FUNCTION_BLOCK FB_Snapshot		// 이번 스캔의 장비 상태를 한 번에 복사. 이후 단계는 이 사본만 읽는다
VAR_IN_OUT
	iq_aipPcs		: ARRAY[1..GVL_PARAM.PCS_COUNT] OF I_Pcs;
	iq_aipBms		: ARRAY[1..GVL_PARAM.BMS_COUNT] OF I_Bms;
	iq_aipMeter		: ARRAY[1..GVL_PARAM.METER_COUNT] OF I_Meter;
END_VAR
VAR_IN_OUT CONSTANT
	iq_astUnitCfg	: ARRAY[1..GVL_PARAM.UNIT_COUNT] OF ST_UnitCfg;
END_VAR
VAR_OUTPUT
	q_astUnit		: ARRAY[1..GVL_PARAM.UNIT_COUNT] OF ST_UnitState;
	q_astBms		: ARRAY[1..GVL_PARAM.BMS_COUNT] OF ST_BatState;
	q_astMeter		: ARRAY[1..GVL_PARAM.METER_COUNT] OF ST_MeterState;
END_VAR
VAR_TEMP
	i				: UINT;
	nPcs			: UINT;
	stNoUnit		: ST_UnitState;		// 빈 칸: 통신 없음, 상태 Unknown
	stNoBms			: ST_BatState;
	stNoMeter		: ST_MeterState;
	k				: UINT;		// [결함 9 수정 2026-11-03: 추가]
END_VAR

// 유닛: 구성표의 PCS 번호·PCS 안 번호로 찾음
FOR i := 1 TO GVL_PARAM.UNIT_COUNT DO
	nPcs := iq_astUnitCfg[i].nPcs;
	IF nPcs >= 1 AND nPcs <= GVL_PARAM.PCS_COUNT AND_THEN iq_aipPcs[nPcs] <> 0 THEN
		q_astUnit[i] := iq_aipPcs[nPcs].M_GetUnitState(iq_astUnitCfg[i].nSub);
		q_astUnit[i].stP := M_FixVal(q_astUnit[i].stP);	// [결함 9 수정 2026-11-03: NaN·무한대 → 0·무효]
		q_astUnit[i].stQ := M_FixVal(q_astUnit[i].stQ);
	ELSE
		q_astUnit[i] := stNoUnit;
	END_IF
END_FOR

FOR i := 1 TO GVL_PARAM.BMS_COUNT DO
	IF iq_aipBms[i] <> 0 THEN
		q_astBms[i] := iq_aipBms[i].BatState;
		q_astBms[i].stSoc := M_FixVal(q_astBms[i].stSoc);	// [결함 9 수정 2026-11-03: NaN·무한대 → 0·무효, 한도는 0]
		q_astBms[i].stSoh := M_FixVal(q_astBms[i].stSoh);
		IF NOT F_CmdOk(q_astBms[i].fPChgMax, 0.0) THEN q_astBms[i].fPChgMax := 0.0; END_IF
		IF NOT F_CmdOk(q_astBms[i].fPDisMax, 0.0) THEN q_astBms[i].fPDisMax := 0.0; END_IF
	ELSE
		q_astBms[i] := stNoBms;
	END_IF
END_FOR

FOR i := 1 TO GVL_PARAM.METER_COUNT DO
	IF iq_aipMeter[i] <> 0 THEN
		q_astMeter[i] := iq_aipMeter[i].MeterState;
		q_astMeter[i].stP := M_FixVal(q_astMeter[i].stP);	// [결함 9 수정 2026-11-03: NaN·무한대 → 0·무효]
		q_astMeter[i].stQ := M_FixVal(q_astMeter[i].stQ);
		q_astMeter[i].stV := M_FixVal(q_astMeter[i].stV);
		FOR k := 1 TO 3 DO
			q_astMeter[i].astV[k] := M_FixVal(q_astMeter[i].astV[k]);
		END_FOR
		q_astMeter[i].stF := M_FixVal(q_astMeter[i].stF);
	ELSE
		q_astMeter[i] := stNoMeter;
	END_IF
END_FOR

METHOD PRIVATE M_FixVal : ST_Val		// 장비 값이 NaN·무한대면 0·무효로 (뒤 계산·비교에 퍼지지 않게). [결함 9 수정 2026-11-03: 추가]
VAR_INPUT
	i_stVal	: ST_Val;
END_VAR
M_FixVal := i_stVal;
IF NOT F_CmdOk(i_stVal.fValue, 0.0) THEN
	M_FixVal.fValue	:= 0.0;
	M_FixVal.bValid	:= FALSE;
END_IF
END_METHOD

END_FUNCTION_BLOCK

(* stored: Version 1.1.0.1, ProductVersion 3.1.4024.15
   POU FB_Snapshot: Id {d02a9ab3-96f3-42df-abd5-45c4e6aa5900}, SpecialFunc None
   Method M_FixVal: Id {4e0b5a6d-0b73-4385-ab44-5cc6792219b1} *)
